//---------------------------------------------------------------------------------------------------------------
//
//  HAUD 2026.11.07
//
//  - TowerControl - fb_DisposableHeros
//
//    - this class is nothing more than the handshake sequence and a timer
//
//    - the station bitmask is written for each production cycle
//      - ticketing involves a DistributorByTicket and its companion ProcessByTicket
//      - this mock up takes care of both tickets.
//        - Why do you need to send 2 tickets?
//          - Distributor and Process instance do not know each other (and this is on purpose to keep things loose and avoid thight coupling by design)
//            --> sending tickets should be done from one place only, so a Distributor sending a ticket internally to its Process would break that rule.
//            --> The Ticket transports the information about where the movers were sent to
//              --> The Process now needs to be told which stations to activate, the rest is ruled by the bitmask from the ticket. 
//
//    - top level transport abstractions are handshaked here:
//    --------------------------------------------
//    - top level transport abstractions
//      - Instances contain the required transport logic
//      - Instances control their assigned ProcessCollector
//      - Instances are controlled in timer based application
//
//
//---------------------------------------------------------------------------------------------------------------
FUNCTION_BLOCK fb_DisposableHeros // Soldier boy, made of clay, now an empty shell
VAR_INPUT
  Start         : BOOL;           // Back to the front
  DwellTime     : TIME;           // Sounding of the clock that ticks
  StationMask   : T_PROCESS;      // molded day by day
END_VAR
VAR
  // process index
  _nProcess               : E_INSTANCE; // whoami
  _nProcessConnect        : e_instance; // to whom am I connected? this is an idea to manage the two tickets for Distributor and Process
  _nProcessConnectTarget  : e_instance; // what is the target of the process to whom I am connected

  _stInstanceCtrl         : REFERENCE TO ARRAY[1..MAX_PROCESS] OF ST_INSTANCE_CTRL;
  _stInstanceState        : REFERENCE TO ARRAY[1..MAX_PROCESS] OF ST_INSTANCE_STATE;

  {attribute 'displaymode':='bin'}
  _wActivateStation       : T_PROCESS;
  _stProcessData          : ST_PROCESS_DATA;

  _ItfTicketList          : I_Process_LinkedList;
  _WriteResult            : ST_PROCESS_LIST_RESULT;

  _nState                 : UINT;
  _tonProcess             : Tc2_Standard.TON;

  _nStationCount          : UINT;

  _nTicketCount           : UDINT;  // since this is a mock up, there is no-one to clean this up
  _nTicketCountLimit      : UDINT;  // if <> 0 --> limit is active

  _MessageLevel           : E_MessageType := E_MessageType.eMessageInfo;
  _stMsg                  : ST_Message;

  _tdx                    : UINT;
  _bRandomize             : BOOL;   // irregular station bitmasks testing
  _eResult                : E_PROGRESS;

  _nLoadCaseOld,
  _nLoadCase              : UINT := 1;

  _nMaskZeroCount         : uint;
END_VAR

//---------------------------------------------------------------------------------------------------------------
//---------------------------------------------------------------------------------------------------------------
// CHECK() ??
// !! this is mock up code, there is no check
//
//---------------------------------------------------------------------------------------------------------------
//---------------------------------------------------------------------------------------------------------------
IF NOT Start THEN _nState   := 0; END_IF
//---------------------------------------------------------------------------------------------------------------
CASE _nState OF
  0:
    IF Start
    THEN
      _nState               := 10;
    END_IF

  10:
    CASE _stInstanceState[_nProcess].ProcessState
    OF
      E_INSTANCE_STATE.DISABLED:
        _stInstanceCtrl[_nProcess].Cmd        := E_INSTANCE_CMD.ENABLE;
        IF (_nProcessConnect > e_instance.INSTANCE_NULL)
        THEN
          memset(ADR(_stProcessData), 0, SIZEOF(_stProcessData));
          _nState                             := 20;
          _wActivateStation                   := StationMask; // this one is important, must be double checked before sending
          _nStationCount                      := _stInstanceState[_nProcessConnect].StationCount;
        END_IF

      E_INSTANCE_STATE.ENABLED:
        CASE _stInstanceState[_nProcess].ProcessProgress
        OF
          E_PROGRESS.PROGRESS_OCCUPIED:       // allow infeed movement
            _stInstanceCtrl[_nProcess].Cmd    := E_INSTANCE_CMD.PROCEED;
        END_CASE

      E_INSTANCE_STATE.WORKING:               // this is for the ProcessByTicket standstill handshake
        CASE _stInstanceState[_nProcess].ProcessProgress
        OF
          E_PROGRESS.PROGRESS_BUSY:           // now every mover has arrived.
            _tonProcess(IN := FALSE, 
                        PT := DwellTime);

            _stInstanceCtrl[_nProcess].Cmd    := E_INSTANCE_CMD.WORK;

          E_PROGRESS.PROGRESS_OCCUPIED:       // time is fleeting
            _tonProcess(IN := TRUE, 
                        PT := DwellTime);

            IF (_tonProcess.Q)
            THEN
              memset(ADR(_stProcessData), 0, SIZEOF(_stProcessData));
              _stInstanceCtrl[_nProcess].Cmd  := E_INSTANCE_CMD.FINISH;
            END_IF
        END_CASE

      E_INSTANCE_STATE.FINISH:                // madness takes its toll
        CASE _stInstanceState[_nProcess].ProcessProgress
        OF
          E_PROGRESS.PROGRESS_DONE:
            _tonProcess(IN := FALSE, 
                        PT := DwellTime);

            _stInstanceCtrl[_nProcess].Cmd    := E_INSTANCE_CMD.DISABLE;

            IF (_nProcessConnect > e_instance.INSTANCE_NULL)
            THEN
              memset(ADR(_stProcessData), 0, SIZEOF(_stProcessData));
              _nState                         := 30;
              _wActivateStation               := StationMask; // this one is important, must be double checked before sending
            END_IF
        END_CASE
    END_CASE
END_CASE
CASE _nState 
OF
  20:
    _nState                                   :=  10;
    TruncMask();

  30:
    IF NOT (_bRandomize)
    THEN
      _nState                                 := 100;
      TruncMask();
    ELSE
      _nState                                 :=  90;
      _eResult                                := ListData(FALSE);
    END_IF
END_CASE
CASE _nState 
OF
  90:
    _eResult                                  := ListData(TRUE);
    IF (_eResult = E_PROGRESS.PROGRESS_DONE)
    THEN
      _nState                                 := 100;
      TruncMask();
    END_IF
END_CASE
CASE _nState 
OF
 100:
  IF NOT (_stProcessData.wTarget > 0)
  THEN
    _nMaskZeroCount                           := _nMaskZeroCount + 1;
    _nTicketCount                             := _nTicketCount + 1;
    _nState                                   := 30;
  ELSE
    IF (_ItfTicketList.Free > 1)
    THEN
      _nState                                 := 101;
    END_IF
  END_IF
END_CASE
CASE _nState 
OF
  101:
    //-----------------------------------------------------------------------------  
    // the tickets
    //-----------------------------------------------------------------------------
    // first send the ticket to the Distributor
    _WriteResult                          := _ItfTicketList.AddTailValue(_stProcessData);
    // second write the ticket for the Process
    _stProcessData.nProcessId             := _nProcessConnect;
    _stProcessData.nTargetId              := _nProcessConnectTarget;
    // third send the ticket to the Process
    _WriteResult                          := _ItfTicketList.AddTailValue(_stProcessData);
    //-----------------------------------------------------------------------------
    _nTicketCount                         := _nTicketCount + 1;
    //-----------------------------------------------------------------------------
    _nState                               := 1000;
END_CASE
CASE _nState 
OF
  1000:
    IF NOT (_nTicketCountLimit > 0)
    THEN
      _nState                             := 0;
    ELSE
      IF (_nTicketCount < _nTicketCountLimit)
      THEN
        _nState                           := 0;
      END_IF
    END_IF
END_CASE

METHOD PUBLIC BitGet : BOOL
VAR_INPUT
  inVal   : T_PROCESS;
  bitNo   : DINT;
END_VAR
VAR
  wConst : T_PROCESS := 1;
END_VAR
IF ( inVal AND SHL( wConst,TO_SINT(bitNo) MOD TO_INT(SIZEOF(T_PROCESS)*8) ) ) > 0
THEN
  BitGet := TRUE;
ELSE
  BitGet := FALSE;
END_IF
END_METHOD

PROPERTY BitmaskRandom : bool
GET
BitmaskRandom := _bRandomize;
END_GET
SET
_bRandomize := BitmaskRandom;
END_SET
END_PROPERTY

METHOD PUBLIC BitSet : T_PROCESS
VAR_INPUT
  inVal   : T_PROCESS;
  bitNo   : DINT;
END_VAR
VAR
  wConst  : T_PROCESS := 1;
END_VAR
BitSet := inVal OR SHL( wConst,TO_SINT(bitNo) MOD TO_INT(SIZEOF(T_PROCESS)*8) );
END_METHOD

PROPERTY InstanceCtrl : REFERENCE TO ARRAY[1..MAX_PROCESS] OF ST_INSTANCE_CTRL
SET
_stInstanceCtrl ref= InstanceCtrl;
END_SET
END_PROPERTY

PROPERTY InstanceState : REFERENCE TO ARRAY[1..MAX_PROCESS] OF ST_INSTANCE_STATE
SET
_stInstanceState ref= InstanceState;
END_SET
END_PROPERTY

METHOD ListData   : E_PROGRESS  // simulates data entry from transfersystem into BUFFER_INFEED linked list
VAR_INPUT
  Execute         : BOOL;
END_VAR
VAR_INST
  _nBit,
  _nExp           : BYTE;
  _nMod           : UINT := 5;

  _eStateProgress,
  _eRslt          : E_PROGRESS;

  _ProcessData    : ST_PROCESS_DATA;

  _nMinListCount  : UDINT := 1;
  _nWaitcountLast,
  _nWaitCount     : UDINT;

  _tMsg           : ST_Message;
END_VAR
//---------------------------------------------------------------------------------------
//---------------------------------------------------------------------------------------
IF NOT Execute THEN _eStateProgress := E_PROGRESS.PROGRESS_INIT; END_IF
//---------------------------------------------------------------------------------------
//---------------------------------------------------------------------------------------
CASE _eStateProgress
OF
   E_PROGRESS.PROGRESS_INIT:
    IF Execute
    THEN
      _eStateProgress         :=  E_PROGRESS.PROGRESS_BUSY;

      IF (_MessageLevel > E_MessageType.eMessageError)
      THEN
        _tMsg.eType           := E_MessageType.eMessageInfo;
        _tMsg.eSubdevice      := e_Subdevice.Application;
        _tMsg.iErrorNumber    := _nTicketCount;
        _tMsg.sText           := concat('ListData.TicketCount: ', TO_STRING(_nTicketCount));
        f_MessageSet(_tMsg);
      END_IF
    END_IF

  E_PROGRESS.PROGRESS_BUSY:
    CASE _nLoadCase
    OF
      0:  // fully loaded
        _eStateProgress       := E_PROGRESS.PROGRESS_CHECK;
        _nLoadCaseOld         := _nLoadCase;

        IF (_MessageLevel > E_MessageType.eMessageError)
        THEN
          _tMsg.eType         := E_MessageType.eMessageInfo;
          _tMsg.eSubdevice    := e_Subdevice.Application;
          _tMsg.iErrorNumber  := _nLoadCase;
          _tMsg.sText         := concat('ListData.Progress: ', TO_STRING(_eStateProgress));
          _tMsg.sText         := concat(_tMsg.sText, ': LoadCase: ');
          _tMsg.sText         := concat(_tMsg.sText, TO_STRING(_nLoadCase));
   
          f_MessageSet(_tMsg);
        END_IF


      1:  // static bits
        _eStateProgress       := E_PROGRESS.PROGRESS_PREPARE;
        _nLoadCaseOld         := _nLoadCase;

        IF (_MessageLevel > E_MessageType.eMessageError)
        THEN
          _tMsg.eType         := E_MessageType.eMessageInfo;
          _tMsg.eSubdevice    := e_Subdevice.Application;
          _tMsg.iErrorNumber  := _nLoadCase;
          _tMsg.sText         := concat('ListData.Progress: ', TO_STRING(_eStateProgress));
          _tMsg.sText         := concat(_tMsg.sText, ': LoadCase: ');
          _tMsg.sText         := concat(_tMsg.sText, TO_STRING(_nLoadCase));
          f_MessageSet(_tMsg);
        END_IF


      2:  // incrementing bits
        _eStateProgress       := E_PROGRESS.PROGRESS_STARTUP;
        _nLoadCaseOld         := _nLoadCase;

        IF (_MessageLevel > E_MessageType.eMessageError)
        THEN
          _tMsg.eType         := E_MessageType.eMessageInfo;
          _tMsg.eSubdevice    := e_Subdevice.Application;
          _tMsg.iErrorNumber  := _nLoadCase;
          _tMsg.sText         := concat('ListData.Progress: ', TO_STRING(_eStateProgress));
          _tMsg.sText         := concat(_tMsg.sText, ': LoadCase: ');
          _tMsg.sText         := concat(_tMsg.sText, TO_STRING(_nLoadCase));
          f_MessageSet(_tMsg);
        END_IF


      99:
        _eStateProgress       := E_PROGRESS.PROGRESS_WORKING;
        _ProcessData.wTarget  := 0;

        IF (_MessageLevel > E_MessageType.eMessageError)
        THEN
          _tMsg.eType          := E_MessageType.eMessageInfo;
          _tMsg.eSubdevice     := e_Subdevice.Application;
          _tMsg.iErrorNumber   := _nLoadCase;
          _tMsg.sText          := concat('sending empty ticket', ': _ProcessData.wTarget: ');
          _tMsg.sText          := concat(_stMsg.sText, f_BitsToString(_ProcessData.wTarget));
          f_MessageSet(_tMsg);
        END_IF
        _nLoadCase            := _nLoadCaseOld;

    ELSE
        _eStateProgress       := E_PROGRESS.PROGRESS_STARTUP;
    END_CASE
    _nWaitCount               := 0; 
END_CASE
//---------------------------------------------------------------------------------------
//---------------------------------------------------------------------------------------
CASE _eStateProgress
OF
  E_PROGRESS.PROGRESS_PREPARE:
    _eStateProgress           := E_PROGRESS.PROGRESS_WORKING;
    _nExp                     := TO_BYTE(_nStationCount);
    _ProcessData.wTarget      := f_To_T_Process(_nExp);

    IF (_nTicketCount MOD _nMod = 0)
    THEN
      _nBit                   := SEL((_nBit>_nExp), _nBit+1, 0);
      _ProcessData.wTarget    := f_BitDel(_ProcessData.wTarget, _nBit);
    END_IF
    IF (_nTicketCount MOD (4) = 0)
    THEN
      _nBit                   := 1;
      _ProcessData.wTarget    := f_BitDel(_ProcessData.wTarget, _nBit);
    END_IF
    IF (_nTicketCount MOD (6) = 0)
    THEN
      _nBit                   := 2;
      _ProcessData.wTarget    := f_BitDel(_ProcessData.wTarget, _nBit);
    END_IF
    IF (_nTicketCount MOD (8) = 0)
    THEN
      _nBit                   := 3;
      _ProcessData.wTarget    := f_BitDel(_ProcessData.wTarget, _nBit);
    END_IF
    IF (_nTicketCount MOD (10) = 0)
    THEN
      _nBit                   := 4;
      _ProcessData.wTarget    := f_BitDel(_ProcessData.wTarget, _nBit);
    END_IF
    IF (_nTicketCount MOD (8) = 0)
    THEN
      _nBit                   := 5;
      _ProcessData.wTarget    := f_BitDel(_ProcessData.wTarget, _nBit);
    END_IF
    IF (_nTicketCount MOD (6) = 0)
    THEN
      _nBit                   := 6;
      _ProcessData.wTarget    := f_BitDel(_ProcessData.wTarget, _nBit);
    END_IF
    IF (_nTicketCount MOD (4) = 0)
    THEN
      _nBit                   := 7;
      _ProcessData.wTarget    := f_BitDel(_ProcessData.wTarget, _nBit);
    END_IF
    IF (_nTicketCount MOD (2) = 0)
    THEN
      _nBit                   := 8;
      _ProcessData.wTarget    := f_BitDel(_ProcessData.wTarget, _nBit);
    END_IF
    IF (_nTicketCount MOD (8) = 0)
    THEN
      _nBit                   := 9;
      _ProcessData.wTarget    := f_BitDel(_ProcessData.wTarget, _nBit);
    END_IF
    IF (_nTicketCount MOD (6) = 0)
    THEN
      _nBit                   := 10;
      _ProcessData.wTarget    := f_BitDel(_ProcessData.wTarget, _nBit);
    END_IF
    IF (_nTicketCount MOD (4) = 0)
    THEN
      _nBit                   := 11;
      _ProcessData.wTarget    := f_BitDel(_ProcessData.wTarget, _nBit);
    END_IF
    IF (_nTicketCount MOD (10) = 0)
    THEN
      _nBit                   := 12;
      _ProcessData.wTarget    := f_BitDel(_ProcessData.wTarget, _nBit);
    END_IF
    IF (_nTicketCount MOD (12) = 0)
    THEN
      _nBit                   := 13;
      _ProcessData.wTarget    := f_BitDel(_ProcessData.wTarget, _nBit);
    END_IF
    IF (_nTicketCount MOD (30) = 0)
    THEN
      _nBit                   := 14;
      _ProcessData.wTarget    := f_BitDel(_ProcessData.wTarget, _nBit);
    END_IF
    IF (_MessageLevel > E_MessageType.eMessageInfo)
    THEN
      _tMsg.eType             := E_MessageType.eMessageInfo;
      _tMsg.eSubdevice        := e_Subdevice.Application;
      _tMsg.iErrorNumber      := _nLoadCase;
      _tMsg.sText             := 'ListData.Progress: ';
      _tMsg.sText             := concat(_tMsg.sText, ': _ProcessData.wTarget: ');
      _tMsg.sText             := concat(_tMsg.sText, f_BitsToString(_ProcessData.wTarget));
      f_MessageSet(_tMsg);
    END_IF
END_CASE
//---------------------------------------------------------------------------------------
//---------------------------------------------------------------------------------------
CASE _eStateProgress
OF
  E_PROGRESS.PROGRESS_STARTUP:
    _eStateProgress           := E_PROGRESS.PROGRESS_WORKING;
    _nExp                     := TO_BYTE(_nStationCount);
    _ProcessData.wTarget      := f_To_T_Process(_nExp);

    IF (_nTicketCount MOD _nMod = 0)
    THEN
      _nBit                   := SEL((_nBit>_nExp), _nBit+1, 0);
      _ProcessData.wTarget    := f_BitDel(_ProcessData.wTarget, _nBit);
    END_IF
    IF (_MessageLevel > E_MessageType.eMessageInfo)
    THEN
      _tMsg.eType             := E_MessageType.eMessageInfo;
      _tMsg.eSubdevice        := e_Subdevice.Application;
      _tMsg.iErrorNumber      := _nLoadCase;
      _tMsg.sText             := 'ListData.Progress: ';
      _tMsg.sText             := concat(_tMsg.sText, ': _ProcessData.wTarget: ');
      _tMsg.sText             := concat(_tMsg.sText, f_BitsToString(_ProcessData.wTarget));
      f_MessageSet(_tMsg);
    END_IF
END_CASE
//---------------------------------------------------------------------------------------
//---------------------------------------------------------------------------------------
CASE _eStateProgress
OF
  E_PROGRESS.PROGRESS_CHECK:
    _eStateProgress           := E_PROGRESS.PROGRESS_WORKING;
    _nExp                     := TO_BYTE(_nStationCount);
    _ProcessData.wTarget      := f_To_T_Process(_nExp);

    IF (_MessageLevel > E_MessageType.eMessageinfo)
    THEN
      _tMsg.eType             := E_MessageType.eMessageInfo;
      _tMsg.eSubdevice        := e_Subdevice.Application;
      _tMsg.iErrorNumber      := _nLoadCase;
      _tMsg.sText             := 'ListData.Progress: ';
      _tMsg.sText             := concat(_tMsg.sText, ': _ProcessData.wTarget: ');
      _tMsg.sText             := concat(_tMsg.sText, f_BitsToString(_ProcessData.wTarget));
      f_MessageSet(_tMsg);
    END_IF
END_CASE
//---------------------------------------------------------------------------------------
//---------------------------------------------------------------------------------------
CASE _eStateProgress
OF
  E_PROGRESS.PROGRESS_WORKING:
    _stProcessData.wTarget    := _ProcessData.wTarget;
    _wActivateStation         := _ProcessData.wTarget;
    _eStateProgress           :=  E_PROGRESS.PROGRESS_DONE;
    IF (_MessageLevel > E_MessageType.eMessageError)
    THEN
      _tMsg.eType             := E_MessageType.eMessageInfo;
      _tMsg.eSubdevice        := e_Subdevice.Application;
      _tMsg.iErrorNumber      := _nLoadCase;
      _tMsg.sText             := 'ListData.Progress: ';
      _tMsg.sText             := concat(_tMsg.sText, ': _wActivateStation: ');
      _tMsg.sText             := concat(_tMsg.sText, f_BitsToString(_ProcessData.wTarget));
      f_MessageSet(_tMsg);
    END_IF
END_CASE
//---------------------------------------------------------------------------------------
//---------------------------------------------------------------------------------------
CASE _eStateProgress
OF
  E_PROGRESS.PROGRESS_OCCUPIED:
    _eStateProgress           :=  E_PROGRESS.PROGRESS_DONE;
END_CASE

ListData                      := _eStateProgress;
END_METHOD

PROPERTY ProcessId : E_INSTANCE
GET
ProcessId := _nProcess;
END_GET
SET
_nProcess := ProcessId;
END_SET
END_PROPERTY

PROPERTY ProcessId_Connect : E_INSTANCE
GET
ProcessId_Connect := _nProcessConnect;
END_GET
SET
_nProcessConnect := ProcessId_Connect;
END_SET
END_PROPERTY

PROPERTY ProcessId_ConnectTarget : E_INSTANCE
GET
ProcessId_ConnectTarget := _nProcessConnectTarget;
END_GET
SET
_nProcessConnectTarget := ProcessId_ConnectTarget;
END_SET
END_PROPERTY

PROPERTY TicketLinkedList : I_Process_LinkedList
SET
_ItfTicketList := TicketLinkedList;
END_SET
END_PROPERTY

METHOD TruncMask : BOOL
VAR_INPUT
END_VAR
// transfer station mask only in the range possible to handle in connected process (StationCount)
_stProcessData.nProcessId                 := _nProcess;
_stProcessData.nTargetId                  := _nProcessConnect;
_stProcessData.wTarget                    := 0;

IF (_nProcessConnect > E_INSTANCE.INSTANCE_NULL) AND
   (_nProcessConnect < E_INSTANCE.INSTANCE_MAX)
THEN
  FOR _tdx := 1 TO _stInstanceState[_nProcessConnect].StationCount
  DO
    IF (BitGet(_wActivateStation, _tdx-1))
    THEN
      _stProcessData.wTarget                := BitSet(_stProcessData.wTarget, _tdx-1);
    END_IF      
  END_FOR
  
  TruncMask := TRUE;
END_IF
END_METHOD

END_FUNCTION_BLOCK

(* stored: Version 1.1.0.1
   POU fb_DisposableHeros: Id {57ff81e0-db35-4988-adb1-755f5d46de47}, SpecialFunc None
   Method BitGet: Id {57c98de9-b3fd-4f7e-920b-502f6210a0a0}
   Property BitmaskRandom: Id {3a95f877-2a5e-4289-9742-41f0517274fd}
   Get Get: Id {19607b5b-25da-455b-b418-a287b5c5ce3c}
   Set Set: Id {4dc908cd-b264-48d9-8bd4-e96a12042123}
   Method BitSet: Id {075d513b-2170-4aca-a2e9-2a16152dac6f}
   Property InstanceCtrl: Id {3363ce1e-638f-4a56-a7d9-502d7b3ac384}
   Set Set: Id {f01b16e3-e7c7-4d66-96b7-a5ce7482bb16}
   Property InstanceState: Id {4aad0611-ac13-4ac9-9913-e5032aa8988a}
   Set Set: Id {d6f80117-bb3a-400d-a886-057ce4f9cae4}
   Method ListData: Id {e0f3ecd8-3034-4b99-ab79-56c0741e0803}
   Property ProcessId: Id {b0d1a924-6241-4335-be39-966d3f9b0719}
   Get Get: Id {4b563e78-35ca-46fa-a429-91bad99e170e}
   Set Set: Id {566aa5ef-d2c9-4a5c-8d5d-3fca3942f3dd}
   Property ProcessId_Connect: Id {abcc06e1-efe7-4aa9-9516-be1588519f38}
   Get Get: Id {b63ddabd-1e94-4d54-b9cd-0e5cfc49b660}
   Set Set: Id {97104ab0-4bc8-47e4-aa6e-413c64ff8466}
   Property ProcessId_ConnectTarget: Id {da385cf2-47a3-4307-bcdb-9af574222ed1}
   Get Get: Id {e9f241da-b82b-4801-b1f0-50eb7bef7352}
   Set Set: Id {95ea77ba-8c13-4f5b-b98e-17a763290a3b}
   Property TicketLinkedList: Id {47e1ba62-2d3b-414e-8705-080e812d120b}
   Set Set: Id {567f8792-66d5-433e-904b-9d5e5e8f13f8}
   Method TruncMask: Id {1e1b7bd6-e3e6-45f2-a35b-d0a434ac7ca6} *)
